TYPE ST_TraceabilityData :
STRUCT
	sName					:STRING(15);
	sValue					:STRING(15);
	sUnit					:STRING(5);
END_STRUCT
END_TYPE

(* stored: Version 1.1.0.1, ProductVersion 3.1.4024.15
   DUT ST_TraceabilityData: Id {9d2302d7-6a8c-4271-83ae-1f022532c8ef} *)
